TYPE ST_VisuPLC_To_PLC :
STRUCT
	lifeBit: BOOL;
	
	RPM_setPoint: REAL;
	
	bPauseTriBlender: BOOL;
	
	bActualComponentDisolving_Done: BOOL;



END_STRUCT
END_TYPE

(* stored: Version 1.1.0.1, ProductVersion 3.1.4024.15
   DUT ST_VisuPLC_To_PLC: Id {02e2d259-713c-4404-b636-e7d4b17005e8} *)
